Fanuc KAREL source: KT00843.KL

PROGRAM KT00843
%NOLOCKGROUP
VAR
  S1: STRING[80]
  S2: STRING[80]
  OUT: REAL
BEGIN
  S1 = 'A'
  S2 = 'B'
  S1 = 'A'
  S2 = 'B'
  OUT = SQRT(S1)
END KT00843
